TYPE "DT_DIGITAL_INPUT_TURBINE"
VERSION : 0.1
   STRUCT
      WICKET_GATE_DISTORSION { S7_SetPoint := 'False'} : "DT_STATUS_SOLO" := ((FALSE, 1, 352), (32000, 32000, 32000), (0, 1, 3), (FALSE, FALSE, 0));
      SPRING_LINK_MONITORING { S7_SetPoint := 'False'} : "DT_STATUS_SOLO" := ((FALSE, 1, 353), (32000, 32000, 32000), (0, 0, 0), (FALSE, FALSE, 0));
      RUNNER_VANES_HEATER_MCB_ON { S7_SetPoint := 'False'} : "DT_STATUS_SOLO" := ((FALSE, 1, 354), (32000, 32000, 32000), (0, 3, 4), (FALSE, FALSE, 0));
      RUNNER_VANES_DRIVE_CONT_OFF { S7_SetPoint := 'False'} : "DT_STATUS_SOLO" := ((FALSE, 1, 355), (32000, 32000, 32000), (0, 1, 4), (FALSE, FALSE, 0));
      RUNNER_VANES_DRIVE_CONT_ON { S7_SetPoint := 'False'} : "DT_STATUS_SOLO" := ((FALSE, 1, 356), (32000, 32000, 32000), (0, 1, 4), (FALSE, FALSE, 0));
      WICKET_GATE_HEATER_MCB_ON { S7_SetPoint := 'False'} : "DT_STATUS_SOLO" := ((FALSE, 1, 357), (32000, 32000, 32000), (0, 3, 4), (FALSE, FALSE, 0));
      RUNNER_VANES_DRIVE_CB_ON { S7_SetPoint := 'False'} : "DT_STATUS_SOLO" := ((FALSE, 1, 358), (32000, 32000, 32000), (0, 3, 4), (FALSE, FALSE, 0));
      WICKET_GATE_DRIVE_CB_ON { S7_SetPoint := 'False'} : "DT_STATUS_SOLO" := ((FALSE, 1, 359), (32000, 32000, 32000), (0, 3, 4), (FALSE, FALSE, 0));
      WICKET_GATE_DRIVE_CONT_OFF { S7_SetPoint := 'False'} : "DT_STATUS_SOLO" := ((FALSE, 1, 360), (32000, 32000, 32000), (0, 1, 4), (FALSE, FALSE, 0));
      WICKET_GATE_DRIVE_CONT_ON { S7_SetPoint := 'False'} : "DT_STATUS_SOLO" := ((FALSE, 1, 361), (32000, 32000, 32000), (0, 1, 4), (FALSE, FALSE, 0));
      WICKET_GATE_HEATER_CONT_ON { S7_SetPoint := 'False'} : "DT_STATUS_SOLO" := ((FALSE, 1, 362), (32000, 32000, 32000), (0, 1, 4), (FALSE, FALSE, 0));
      OVERSPEED_PROT_TRIP_TURB { S7_SetPoint := 'False'} : "DT_STATUS_SOLO" := ((FALSE, 1, 363), (32000, 32000, 32000), (0, 1, 3), (FALSE, FALSE, 0));
      WICKET_GATE_TORQUE_SWITCH_C { S7_SetPoint := 'False'} : "DT_STATUS_SOLO" := ((FALSE, 1, 364), (32000, 32000, 32000), (0, 1, 3), (FALSE, FALSE, 0));
      WICKET_GATE_TORQUE_SWITCH_O { S7_SetPoint := 'False'} : "DT_STATUS_SOLO" := ((FALSE, 1, 365), (32000, 32000, 32000), (0, 1, 3), (FALSE, FALSE, 0));
      WICKET_GATE_LIMIT_SWITCH_C { S7_SetPoint := 'False'} : "DT_STATUS_SOLO" := ((FALSE, 1, 366), (32000, 32000, 32000), (0, 1, 3), (FALSE, FALSE, 0));
      WICKET_GATE_LIMIT_SWITCH_O { S7_SetPoint := 'False'} : "DT_STATUS_SOLO" := ((FALSE, 1, 367), (32000, 32000, 32000), (0, 1, 3), (FALSE, FALSE, 0));
      RUNNER_VANES_TORQUE_SWITCH_C { S7_SetPoint := 'False'} : "DT_STATUS_SOLO" := ((FALSE, 1, 368), (32000, 32000, 32000), (0, 1, 3), (FALSE, FALSE, 0));
      RUNNER_VANES_TORQUE_SWITCH_O { S7_SetPoint := 'False'} : "DT_STATUS_SOLO" := ((FALSE, 1, 369), (32000, 32000, 32000), (0, 1, 3), (FALSE, FALSE, 0));
      RUNNER_VANES_LIMIT_SWITCH_C { S7_SetPoint := 'False'} : "DT_STATUS_SOLO" := ((FALSE, 1, 370), (32000, 32000, 32000), (0, 1, 3), (FALSE, FALSE, 0));
      RUNNER_VANES_LIMIT_SWITCH_O { S7_SetPoint := 'False'} : "DT_STATUS_SOLO" := ((FALSE, 1, 371), (32000, 32000, 32000), (0, 1, 3), (FALSE, FALSE, 0));
      RUNNER_VANES_THERMOSWITCH { S7_SetPoint := 'False'} : "DT_STATUS_SOLO" := ((FALSE, 1, 372), (32000, 32000, 32000), (0, 1, 3), (FALSE, FALSE, 0));
      SPARE_373 { S7_SetPoint := 'False'} : "DT_STATUS_SOLO" := ((FALSE, 1, 373), (32000, 32000, 32000), (0, 0, 0), (FALSE, FALSE, 0));
      SPARE_374 { S7_SetPoint := 'False'} : "DT_STATUS_SOLO" := ((FALSE, 1, 374), (32000, 32000, 32000), (0, 0, 0), (FALSE, FALSE, 0));
      SPARE_375 { S7_SetPoint := 'False'} : "DT_STATUS_SOLO" := ((FALSE, 1, 375), (32000, 32000, 32000), (0, 0, 0), (FALSE, FALSE, 0));
      SPARE_376 { S7_SetPoint := 'False'} : "DT_STATUS_SOLO" := ((FALSE, 1, 376), (32000, 32000, 32000), (0, 0, 0), (FALSE, FALSE, 0));
      SPARE_377 { S7_SetPoint := 'False'} : "DT_STATUS_SOLO" := ((FALSE, 1, 377), (32000, 32000, 32000), (0, 0, 0), (FALSE, FALSE, 0));
      SPARE_378 { S7_SetPoint := 'False'} : "DT_STATUS_SOLO" := ((FALSE, 1, 378), (32000, 32000, 32000), (0, 0, 0), (FALSE, FALSE, 0));
      SPARE_379 { S7_SetPoint := 'False'} : "DT_STATUS_SOLO" := ((FALSE, 1, 379), (32000, 32000, 32000), (0, 0, 0), (FALSE, FALSE, 0));
      SPARE_380 { S7_SetPoint := 'False'} : "DT_STATUS_SOLO" := ((FALSE, 1, 380), (32000, 32000, 32000), (0, 0, 0), (FALSE, FALSE, 0));
      SPARE_381 { S7_SetPoint := 'False'} : "DT_STATUS_SOLO" := ((FALSE, 1, 381), (32000, 32000, 32000), (0, 0, 0), (FALSE, FALSE, 0));
      SPARE_382 { S7_SetPoint := 'False'} : "DT_STATUS_SOLO" := ((FALSE, 1, 382), (32000, 32000, 32000), (0, 0, 0), (FALSE, FALSE, 0));
      SPARE_383 { S7_SetPoint := 'False'} : "DT_STATUS_SOLO" := ((FALSE, 1, 383), (32000, 32000, 32000), (0, 0, 0), (FALSE, FALSE, 0));
   END_STRUCT;

END_TYPE

